(* IEC 61131-3 sources: codesys-framework/txt/application/ToDo/Utils/Moving Average/FB_MovingAverage, 6 files *)

(* ---- AddValue.method.st ---- *)
METHOD AddValue
VAR_INPUT
	lrValue 	: LREAL;
END_VAR

// --- BEGIN IMPLEMENTATION ---

_iInsertIndex := _iInsertIndex + 1;

IF _iInsertIndex > _iNbrOfItems THEN
	_iInsertIndex := 1;
END_IF

IF _iNbrOfItemsInList < _iNbrOfItems THEN
	_iNbrOfItemsInList := _iNbrOfItemsInList + 1;
END_IF

_alrValues[_iInsertIndex] := lrValue;

(* ---- CalculateAverage.method.st ---- *)
METHOD PROTECTED  CalculateAverage
VAR_INPUT
	alrValues 	: ARRAY[1..cMaxNbrOfEntries] OF LREAL;
END_VAR
VAR
	lrTotal 	: LREAL;
	lrAverage 	: LREAL;
	i 			: UINT;
END_VAR

// --- BEGIN IMPLEMENTATION ---

lrTotal := 0;
lrAverage := 0;

FOR i := 1 TO _iNbrOfItems DO
	lrTotal := lrTotal + alrValues[i];
END_FOR

IF _iNbrOfItemsInList > 0 THEN
	lrAverage := lrTotal / _iNbrOfItemsInList;
ELSE
	lrAverage := 0;
END_IF

_lrAverage := lrAverage;

(* ---- CheckNumberOfItems.method.st ---- *)
METHOD PRIVATE CheckNumberOfItems
VAR_INPUT
END_VAR

// --- BEGIN IMPLEMENTATION ---

_iNbrOfItems := _scSysPar.iNbrOfItemsForAverage;

IF _iNbrOfItems <= 0 THEN
	_iNbrOfItems := 10;
END_IF

IF _iNbrOfItems > cMaxNbrOfEntries THEN
	_iNbrOfItems := cMaxNbrOfEntries;
END_IF

(* ---- GetAverage.method.st ---- *)
METHOD GetAverage : lREAL
VAR_INPUT
END_VAR

// --- BEGIN IMPLEMENTATION ---

GetAverage := _lrAverage;

(* ---- Reset.method.st ---- *)
METHOD Reset
VAR_INPUT
END_VAR
VAR
	i 	: UINT;
END_VAR

// --- BEGIN IMPLEMENTATION ---

FOR i := 1 TO cMaxNbrOfEntries DO
	_alrValues[i] := 0;
END_FOR

_lrAverage := 0;
_iInsertIndex := 0;
_iNbrOfItemsInList := 0;

(* ---- SysPar.prop.st ---- *)
PROPERTY SysPar : SC_SystemParametersMovingAverage

// --- BEGIN IMPLEMENTATION ---

// ----------- SET -----------
VAR
END_VAR

// -- BEGIN IMPLEMENTATION SET --
_scSysPar := SysPar;
